(* IEC 61131-3 sources: plc-vscode/tests/st/test-ready/rusty/tests/lit/single/init, 58 files *)

(* ---- array_alias_struct_init.st ---- *)
// RUN: (%COMPILE %s && %RUN) | %CHECK %s

// Verify that array type aliases with struct initializers produce correct runtime values.
TYPE SomeStruct : STRUCT
    field4 : USINT;
END_STRUCT
END_TYPE

TYPE SomeArray : ARRAY[1..2] OF SomeStruct; END_TYPE
TYPE MySomeArrayWInit : SomeArray := [(field4 := 1), (field4 := 2)]; END_TYPE

VAR_GLOBAL
    g_arr : MySomeArrayWInit;
END_VAR

FUNCTION main : DINT
VAR
    local_arr : MySomeArrayWInit;
END_VAR
    // Global instance should carry the type-level initializer
    printf('%d$N', g_arr[1].field4);   // CHECK: 1
    printf('%d$N', g_arr[2].field4);   // CHECK: 2

    // Local instance should also be initialized via the type ctor
    printf('%d$N', local_arr[1].field4);  // CHECK: 1
    printf('%d$N', local_arr[2].field4);  // CHECK: 2
    main := 0;
END_FUNCTION

(* ---- array_constant_indirect_type_init.st ---- *)
// RUN: (%COMPILE %s && %RUN) | %CHECK %s

TYPE IntArrayBase : ARRAY[1..3] OF DINT := [11, 22, 33]; END_TYPE
TYPE IntArrayAlias : IntArrayBase; END_TYPE
TYPE IntArrayAlias2 : IntArrayAlias; END_TYPE

VAR_GLOBAL CONSTANT
    g_base : IntArrayBase;
    g_alias : IntArrayAlias;
    g_alias2 : IntArrayAlias2;
END_VAR

FUNCTION main : DINT
    printf('g_base=%d,%d,%d$N', g_base[1], g_base[2], g_base[3]); // CHECK: g_base=11,22,33
    printf('g_alias=%d,%d,%d$N', g_alias[1], g_alias[2], g_alias[3]); // CHECK: g_alias=11,22,33
    printf('g_alias2=%d,%d,%d$N', g_alias2[1], g_alias2[2], g_alias2[3]); // CHECK: g_alias2=11,22,33

    main := 0;
END_FUNCTION

(* ---- array_external_type_init.st ---- *)
// RUN: (%COMPILE %s && %RUN) | %CHECK %s

// Verify that arrays with type-level initializers work correctly
// when declared in external blocks.
TYPE tarr : ARRAY[0..4] OF DINT := [5(77)]; END_TYPE

VAR_GLOBAL
    g_arr : tarr;
END_VAR

FUNCTION main : DINT
VAR
    local_arr : tarr;
END_VAR
    // Global instance should be initialized by the global ctor
    printf('%d$N', g_arr[0]);   // CHECK: 77
    printf('%d$N', g_arr[4]);   // CHECK: 77

    // Local instance should also be initialized via the type ctor
    printf('%d$N', local_arr[0]);  // CHECK: 77
    printf('%d$N', local_arr[4]);  // CHECK: 77
    main := 0;
END_FUNCTION

(* ---- array_multiplied_large.st ---- *)
// RUN: (%COMPILE %s && %RUN) | %CHECK %s
TYPE tarr : ARRAY[0..9999] OF DINT := [10000(7)]; END_TYPE

FUNCTION main : DINT
VAR
    arr : tarr;
END_VAR
    // Spot-check first, middle, and last elements
    printf('%d$N', arr[0]);     // CHECK: 7
    printf('%d$N', arr[4999]);  // CHECK: 7
    printf('%d$N', arr[9999]);  // CHECK: 7
    main := 0;
END_FUNCTION

(* ---- array_multiplied_mixed_init.st ---- *)
// RUN: (%COMPILE %s && %RUN) | %CHECK %s
TYPE tarr : ARRAY[0..9] OF DINT := [5(10), 3(20), 99, 100]; END_TYPE

FUNCTION main : DINT
VAR
    arr : tarr;
END_VAR
    // First segment: indices 0..4 should be 10
    printf('%d$N', arr[0]);  // CHECK: 10
    printf('%d$N', arr[4]);  // CHECK: 10
    // Second segment: indices 5..7 should be 20
    printf('%d$N', arr[5]);  // CHECK: 20
    printf('%d$N', arr[7]);  // CHECK: 20
    // Individual values at indices 8 and 9
    printf('%d$N', arr[8]);  // CHECK: 99
    printf('%d$N', arr[9]);  // CHECK: 100
    main := 0;
END_FUNCTION

(* ---- array_multiplied_nonzero_offset.st ---- *)
// RUN: (%COMPILE %s && %RUN) | %CHECK %s
TYPE tarr : ARRAY[10..19] OF DINT := [10(77)]; END_TYPE

FUNCTION main : DINT
VAR
    arr : tarr;
END_VAR
    printf('%d$N', arr[10]);  // CHECK: 77
    printf('%d$N', arr[14]);  // CHECK: 77
    printf('%d$N', arr[19]);  // CHECK: 77
    main := 0;
END_FUNCTION

(* ---- array_multiplied_partial_init.st ---- *)
// RUN: (%COMPILE %s && %RUN) | %CHECK %s
TYPE tarr : ARRAY[0..9] OF DINT := [5(42)]; END_TYPE

FUNCTION main : DINT
VAR
    arr : tarr;
END_VAR
    // First 5 elements should be 42
    printf('%d$N', arr[0]);  // CHECK: 42
    printf('%d$N', arr[4]);  // CHECK: 42
    // Remaining elements should be 0 (default)
    printf('%d$N', arr[5]);  // CHECK: 0
    printf('%d$N', arr[9]);  // CHECK: 0
    main := 0;
END_FUNCTION

(* ---- array_multiplied_struct_elements.st ---- *)
// RUN: (%COMPILE %s && %RUN) | %CHECK %s
TYPE MyStruct : STRUCT
    a : DINT;
    b : DINT;
END_STRUCT END_TYPE

FUNCTION main : DINT
VAR
    arr : ARRAY[0..2] OF MyStruct := [3((a := 5, b := 10))];
END_VAR
    printf('%d %d$N', arr[0].a, arr[0].b);  // CHECK: 5 10
    printf('%d %d$N', arr[1].a, arr[1].b);  // CHECK: 5 10
    printf('%d %d$N', arr[2].a, arr[2].b);  // CHECK: 5 10
    main := 0;
END_FUNCTION

(* ---- array_multiplied_type_init.st ---- *)
// RUN: (%COMPILE %s && %RUN) | %CHECK %s
TYPE tarr : ARRAY[0..99] OF DINT := [100(42)]; END_TYPE

FUNCTION main : DINT
VAR
    arr : tarr;
END_VAR
    // Check first, middle, and last elements
    printf('%d$N', arr[0]);   // CHECK: 42
    printf('%d$N', arr[49]);  // CHECK: 42
    printf('%d$N', arr[99]);  // CHECK: 42
    main := 0;
END_FUNCTION

(* ---- array_of_structs_init.st ---- *)
// RUN: (%COMPILE %s && %RUN) | %CHECK %s

TYPE Point : STRUCT
    x : DINT;
    y : DINT;
END_STRUCT END_TYPE

FUNCTION main : DINT
    VAR
        points : ARRAY[0..1] OF Point := [(x := 1, y := 2), (x := 3, y := 4)];
    END_VAR

    // CHECK: 1
    printf('%d$N', points[0].x);

    // CHECK: 2
    printf('%d$N', points[0].y);

    // CHECK: 3
    printf('%d$N', points[1].x);

    // CHECK: 4
    printf('%d$N', points[1].y);
END_FUNCTION

(* ---- global_nested_struct_with_default_and_override_refs.st ---- *)
// RUN: (%COMPILE %s && %RUN) | %CHECK %s
VAR_GLOBAL
    globalValueA: DINT := 5;
    globalValueB: DINT := 10;
    globalValueC: DINT := 15;

    globalStructOne: StructA;
    globalStructTwo: StructA := (value := REF(globalValueA), instanceB := (value := REF(globalValueB), instanceC := (value := REF(globalValueC))));
END_VAR

TYPE StructA:
    STRUCT
        value: REF_TO DINT := REF(globalValueC);
        instanceB: StructB;
    END_STRUCT
END_TYPE

TYPE StructB:
    STRUCT
        value: REF_TO DINT := REF(globalValueA);
        instanceC: StructC;
    END_STRUCT
END_TYPE

TYPE StructC:
    STRUCT
        value: REF_TO DINT := REF(globalValueB);
    END_STRUCT
END_TYPE

FUNCTION main
    printf('%d$N', globalStructOne.value^); // CHECK: 15
    printf('%d$N', globalStructOne.instanceB.value^); // CHECK: 5
    printf('%d$N', globalStructOne.instanceB.instanceC.value^); // CHECK: 10

    printf('%d$N', globalStructTwo.value^); // CHECK: 5
    printf('%d$N', globalStructTwo.instanceB.value^); // CHECK: 10
    printf('%d$N', globalStructTwo.instanceB.instanceC.value^); // CHECK: 15
END_FUNCTION

(* ---- global_nested_struct_with_mixed_ref_assignments.st ---- *)
// RUN: (%COMPILE %s && %RUN) | %CHECK %s
VAR_GLOBAL
    globalOne: DINT := 1;
    globalTwo: DINT := 2;
    globalThree: DINT := 3;
    globalFour: DINT := 4;
    globalFive: DINT := 5;
    globalSix: DINT := 6;
    globalSeven: DINT := 7;
    globalEight: DINT := 8;
    globalNine: DINT := 9;

    globalA: MyStruct2 := (a := (c := REF(globalFive), b := REF(globalSeven)), b := (a := REF(globalThree), b := REF(globalTwo)));
    globalB: MyStruct2 := (b := (a := REF(globalNine)));
END_VAR

TYPE MyStruct2: STRUCT
    a: MyStruct := (a := REF(globalFive), b := REF(globalFour));
    b: MyStruct := (c := REF(globalSeven));
END_STRUCT
END_TYPE

TYPE MyStruct: STRUCT
    a: REF_TO DINT := REF(globalOne);
    b: REF_TO DINT := REF(globalTwo);
    c: REF_TO DINT := REF(globalThree);
END_STRUCT
END_TYPE

FUNCTION main
    printf('%d$N', globalA.a.a^); // CHECK: 5
    printf('%d$N', globalA.a.b^); // CHECK: 7
    printf('%d$N', globalA.a.c^); // CHECK: 5
    printf('%d$N', globalA.b.a^); // CHECK: 3
    printf('%d$N', globalA.b.b^); // CHECK: 2
    printf('%d$N', globalA.b.c^); // CHECK: 7

    printf('%d$N', globalB.b.a^); // CHECK: 9
    printf('%d$N', globalB.b.b^); // CHECK: 2
    printf('%d$N', globalB.b.c^); // CHECK: 7
END_FUNCTION

(* ---- global_struct_with_partial_nested_initialization.st ---- *)
// RUN: (%COMPILE %s && %RUN) | %CHECK %s
VAR_GLOBAL
    globalFoo: DINT := 15;
    globalBar: DINT := 30;
    globalBar2: DINT := 45;

    globalStructOne: StructA;
    globalStructTwo: StructA := (instanceB := (bar := REF(globalBar2)));
END_VAR

TYPE StructA:
    STRUCT
        instanceB: StructB := (foo := REF(globalFoo));
    END_STRUCT
END_TYPE

TYPE StructB:
    STRUCT
        foo: REF_TO DINT;
        bar: REF_TO DINT := REF(globalBar);
    END_STRUCT
END_TYPE

FUNCTION main
    printf('%d$N', globalStructOne.instanceB.foo^); // CHECK: 15
    printf('%d$N', globalStructOne.instanceB.bar^); // CHECK: 30

    printf('%d$N', globalStructTwo.instanceB.foo^); // CHECK: 15
    printf('%d$N', globalStructTwo.instanceB.bar^); // CHECK: 45
END_FUNCTION

(* ---- local_struct_with_global_ref_initialization.st ---- *)
// RUN: (%COMPILE %s && %RUN) | %CHECK %s
VAR_GLOBAL
    globalVar: DINT := 10;
END_VAR

TYPE Parent:
    STRUCT
        foo: REF_TO DINT;
    END_STRUCT
END_TYPE

TYPE Child:
    STRUCT
        instance: Parent := (foo := REF(globalVar));
    END_STRUCT
END_TYPE

FUNCTION main
    VAR
        localChild: Child;
    END_VAR

    // CHECK: Value: 10
    printf('Value: %d$N', localChild.instance.foo^);
END_FUNCTION

(* ---- struct_array_field_init_from_array.st ---- *)
// Issue #921: Array field initialization from another array in struct literal
// RUN: (%COMPILE %s && %RUN) | %CHECK %s

TYPE myStruct : STRUCT
    var1 : DINT;
    var2 : ARRAY[1..2] OF DINT;
END_STRUCT
END_TYPE

FUNCTION main : DINT
VAR
    arr_init : ARRAY[1..2] OF DINT := [1, 2];
    x : myStruct;
END_VAR
    // Initialize array field from another array (regression for #921)
    x := (var1 := 1, var2 := arr_init);

    printf('v1=%d$N', x.var1); // CHECK: v1=1
    printf('v2_1=%d$N', x.var2[1]); // CHECK: v2_1=1
    printf('v2_2=%d$N', x.var2[2]); // CHECK: v2_2=2

    main := 0;
END_FUNCTION

(* ---- struct_with_array_of_strings_init.st ---- *)
// RUN: (%COMPILE %s && %RUN) | %CHECK %s

TYPE Container : STRUCT
    data : ARRAY[0..2] OF STRING;
END_STRUCT END_TYPE

FUNCTION main : DINT
    VAR
        container : Container := (data := ['one', 'two', 'three']);
    END_VAR

    // CHECK: one
    printf('%s$N', container.data[0]);

    // CHECK: two
    printf('%s$N', container.data[1]);

    // CHECK: three
    printf('%s$N', container.data[2]);
END_FUNCTION

(* ---- struct_with_string_init.st ---- *)
// RUN: (%COMPILE %s && %RUN) | %CHECK %s
TYPE Transaction : STRUCT
    id      : DINT;
    amount  : DINT;
    message : STRING;
END_STRUCT END_TYPE

FUNCTION main : DINT
    VAR
        txn     : Transaction := (id := 1, amount := 5, message := 'whats up');
    END_VAR

    // CHECK: 1
    printf('%d$N', txn.id);

    // CHECK: 5
    printf('%d$N', txn.amount);

    // CHECK: whats up
    printf('%s$N', txn.message);
END_FUNCTION

(* ---- type_alias_initializers.st ---- *)
// RUN: (%COMPILE %s && %RUN) | %CHECK %s

// Comprehensive test for type aliases with initializers (enum, struct, array).
TYPE SomeEnum : (E1, E2, E3); END_TYPE
TYPE MySomeEnumWInit : SomeEnum := E2; END_TYPE

TYPE SomeStruct : STRUCT
    field2 : DINT;
    field3 : BOOL;
    field4 : USINT;
END_STRUCT
END_TYPE
TYPE MySomeStructWInit : SomeStruct := (field3 := FALSE, field2 := 9); END_TYPE

TYPE SomeArray : ARRAY[1..2] OF SomeStruct; END_TYPE
TYPE MySomeArrayWInit : SomeArray := [(field4 := 2), (field4 := 2)]; END_TYPE

// Aliases without custom initializers (should inherit defaults)
TYPE MySomeEnum : SomeEnum; END_TYPE
TYPE MySomeStruct : SomeStruct; END_TYPE
TYPE MySomeArray : SomeArray; END_TYPE

FUNCTION main : DINT
VAR
    e : MySomeEnumWInit;
    s : MySomeStructWInit;
    a : MySomeArrayWInit;
    e_default : MySomeEnum;
    s_default : MySomeStruct;
    a_default : MySomeArray;
END_VAR
    // Enum alias with initializer (E1=0, E2=1)
    printf('%d$N', e);            // CHECK: 1

    // Struct alias with initializer
    printf('%d$N', s.field2);     // CHECK: 9
    printf('%d$N', s.field3);     // CHECK: 0

    // Array alias with struct initializer
    printf('%d$N', a[1].field4);  // CHECK: 2
    printf('%d$N', a[2].field4);  // CHECK: 2

    // Default enum (should be 0 / E1)
    printf('%d$N', e_default);    // CHECK: 0

    // Default struct fields (should be 0)
    printf('%d$N', s_default.field2);  // CHECK: 0

    // Default array element (should be 0)
    printf('%d$N', a_default[1].field4);  // CHECK: 0

    main := 0;
END_FUNCTION

(* ---- typedef_initializer_chain.st ---- *)
// Issue #1522: Typedef initializer chains not propagating values
// RUN: (%COMPILE %s && %RUN) | %CHECK %s

TYPE myStruct: STRUCT
  a : INT;
END_STRUCT
END_TYPE

TYPE mytypedefstruct: myStruct := (a := 3); END_TYPE
TYPE mysubtype: mytypedefstruct; END_TYPE
TYPE mysubtype2: mysubtype; END_TYPE

FUNCTION main : DINT
VAR
    inst: mysubtype2;
END_VAR
    printf('a=%d$N', inst.a); // CHECK: a=3
    main := 0;
END_FUNCTION

(* ---- var_input_defaults_function_array_string.st ---- *)
// RUN: (%COMPILE %s && %RUN) | %CHECK %s

// Test VAR_INPUT defaults with STRING/ARRAY and mixed overrides

TYPE ArrType : ARRAY[1..3] OF DINT;
END_TYPE

FUNCTION test : DINT
VAR_INPUT
    s : STRING := 'abc';
    a : ArrType := [1, 2, 3];
END_VAR
test := a[1] + a[2] + a[3];
printf('s=%s$N', REF(s));
printf('sum=%d$N', test);
END_FUNCTION

FUNCTION main
VAR
    tmp : DINT;
END_VAR
// Defaults (no overrides)
tmp := test();
// CHECK: s=abc
// CHECK: sum=6
printf('case=default$N'); // CHECK: case=default

// Override string only
tmp := test(s := 'xyz');
// CHECK: s=xyz
// CHECK: sum=6
printf('case=string$N'); // CHECK: case=string

// Override array only
tmp := test(a := [4, 5, 6]);
// CHECK: s=abc
// CHECK: sum=15
printf('case=array$N'); // CHECK: case=array

// Override both
tmp := test(s := 'pqr', a := [7, 8, 9]);
// CHECK: s=pqr
// CHECK: sum=24
printf('case=both$N'); // CHECK: case=both
END_FUNCTION

(* ---- var_input_defaults_function_wstring.st ---- *)
// RUN: (%COMPILE %s && %RUN) | %CHECK %s
// Test VAR_INPUT defaults with WSTRING and overrides

TYPE ArrType : ARRAY[1..3] OF DINT;
END_TYPE

FUNCTION test : DINT
VAR_INPUT
    s : STRING := 'abc';
    ws : WSTRING := "def";
    a : ArrType := [1, 2, 3];
    i : DINT := 10;
END_VAR
test := a[1] + a[2] + a[3] + i;
printf('s=%s$N', REF(s));
printf('ws=%s$N', REF(TO_STRING(ws)));
printf('sum=%d$N', test);
END_FUNCTION

FUNCTION main : DINT
    // Case 1: all defaults
    test();
    // CHECK: s=abc
    // CHECK: ws=def
    // CHECK: sum=16

    // Case 2: override one input
    test(s := 'xyz');
    // CHECK: s=xyz
    // CHECK: ws=def
    // CHECK: sum=16

    // Case 3: override WSTRING and array
    test(ws := "uvw", a := [4, 5, 6]);
    // CHECK: s=abc
    // CHECK: ws=uvw
    // CHECK: sum=25

    // Case 4: override all inputs
    test(s := 'qqq', ws := "rst", a := [7, 8, 9], i := 1);
    // CHECK: s=qqq
    // CHECK: ws=rst
    // CHECK: sum=25
END_FUNCTION

(* ---- var_input_ref_defaults_string_array.st ---- *)
// RUN: (%COMPILE %s && %RUN) | %CHECK %s
// Test VAR_INPUT {ref} defaults with STRING/ARRAY and mixed overrides

TYPE ArrType : ARRAY[1..3] OF DINT;
END_TYPE

FUNCTION test : DINT
VAR_INPUT {ref}
    s : STRING;
    a : ArrType;
END_VAR
test := a[1] + a[2] + a[3];
printf('s=%s$N', REF(s));
printf('sum=%d$N', test);
END_FUNCTION

FUNCTION main
VAR
    tmp : DINT;
    s_default : STRING := 'abc';
    s_override : STRING := 'xyz';
    s_both : STRING := 'pqr';
    a_default : ArrType := [1, 2, 3];
    a_override : ArrType := [4, 5, 6];
    a_both : ArrType := [7, 8, 9];
END_VAR
// Defaults (no overrides)
tmp := test(s := s_default, a := a_default);
// CHECK: s=abc
// CHECK: sum=6

// Override string only
tmp := test(s := s_override, a := a_default);
// CHECK: s=xyz
// CHECK: sum=6

// Override array only
tmp := test(s := s_default, a := a_override);
// CHECK: s=abc
// CHECK: sum=15

// Override both
tmp := test(s := s_both, a := a_both);
// CHECK: s=pqr
// CHECK: sum=24
END_FUNCTION

(* ---- array_const_bound_multiplied_real.st ---- *)
// RUN: (%COMPILE %s && %RUN) | %CHECK %s
// Tests that an array with constant-expression bounds and a constant-multiplied
// REAL initializer compiles and runs correctly.

VAR_GLOBAL CONSTANT
    NB_BOOL   : DINT := 12;
    NB_ANALOG : DINT := 2;
END_VAR

FUNCTION main : DINT
VAR
    MAX_TIME_BOOL   : ARRAY [1..NB_BOOL] OF REAL := [(NB_BOOL)(0.0033)];
    MAX_TIME_ANALOG : ARRAY [1..NB_ANALOG] OF REAL := [(NB_ANALOG)(1.5)];
END_VAR
    // Check first, middle, and last elements of MAX_TIME_BOOL
    printf('%.4f$N', MAX_TIME_BOOL[1]);   // CHECK: 0.0033
    printf('%.4f$N', MAX_TIME_BOOL[6]);   // CHECK: 0.0033
    printf('%.4f$N', MAX_TIME_BOOL[12]);  // CHECK: 0.0033

    // Check both elements of MAX_TIME_ANALOG
    printf('%.1f$N', MAX_TIME_ANALOG[1]);  // CHECK: 1.5
    printf('%.1f$N', MAX_TIME_ANALOG[2]);  // CHECK: 1.5

    main := 0;
END_FUNCTION

(* ---- array_const_bound_multiplied_real_global.st ---- *)
// RUN: (%COMPILE %s && %RUN) | %CHECK %s
// Tests that global constant arrays with constant-expression bounds and
// constant-multiplied REAL initializers compile and run correctly.

VAR_GLOBAL CONSTANT
    NB_BOOL       : DINT := 12;
    NB_ANALOG     : DINT := 2;
    MAX_TIME_BOOL   : ARRAY [1..NB_BOOL] OF REAL := [(NB_BOOL)(0.0033)];
    MAX_TIME_ANALOG : ARRAY [1..NB_ANALOG] OF REAL := [(NB_ANALOG)(1.5)];
END_VAR

FUNCTION main : DINT
    // Check first, middle, and last elements of MAX_TIME_BOOL
    printf('%.4f$N', MAX_TIME_BOOL[1]);   // CHECK: 0.0033
    printf('%.4f$N', MAX_TIME_BOOL[6]);   // CHECK: 0.0033
    printf('%.4f$N', MAX_TIME_BOOL[12]);  // CHECK: 0.0033

    // Check both elements of MAX_TIME_ANALOG
    printf('%.1f$N', MAX_TIME_ANALOG[1]);  // CHECK: 1.5
    printf('%.1f$N', MAX_TIME_ANALOG[2]);  // CHECK: 1.5

    main := 0;
END_FUNCTION

(* ---- global_variables.st ---- *)
// RUN: (%COMPILE %s && %RUN) | %CHECK %s
VAR_GLOBAL
    arr : ARRAY[0..3] OF STRING := ['a', 'b', 'c', 'd'];
    alias AT arr : ARRAY[0..3] OF STRING;
END_VAR

FUNCTION main: DINT
    // CHECK: a, b, c, d
    printf('%s, %s, %s, %s$N', REF(alias[0]), REF(alias[1]), REF(alias[2]), REF(alias[3]));
END_FUNCTION

(* ---- ref_initializer_with_array_init.st ---- *)
// RUN: (%COMPILE %s && %RUN) | %CHECK %s

VAR_GLOBAL
    globalString: STRING := 'Global String';
END_VAR

FUNCTION main : DINT
VAR
    localString: REF_TO STRING := REF(globalString);
    arr: ARRAY[1..2] OF DINT := [1, 2];
END_VAR
    printf('ref=%s$N', localString); // CHECK: ref=Global String
    printf('arr1=%d$N', arr[1]); // CHECK: arr1=1
    printf('arr2=%d$N', arr[2]); // CHECK: arr2=2
    main := 0;
END_FUNCTION

(* ---- array_local_const_multiplied.st ---- *)
// RUN: (%COMPILE %s && %RUN) | %CHECK %s
// Tests that a POU-local VAR CONSTANT can be used as the multiplier
// in an array initializer with the [(CONST)(value)] syntax.

FUNCTION main : DINT
VAR CONSTANT
    N     : DINT := 5;
    COUNT : DINT := 3;
END_VAR
VAR
    arr1 : ARRAY [0..4] OF DINT := [(N)(77)];
    arr2 : ARRAY [1..3] OF REAL := [(COUNT)(1.25)];
END_VAR
    printf('%d$N', arr1[0]);  // CHECK: 77
    printf('%d$N', arr1[2]);  // CHECK: 77
    printf('%d$N', arr1[4]);  // CHECK: 77

    printf('%.2f$N', arr2[1]);  // CHECK: 1.25
    printf('%.2f$N', arr2[3]);  // CHECK: 1.25

    main := 0;
END_FUNCTION

(* ---- array_mixed_ref_segments.st ---- *)
// RUN: (%COMPILE %s && %RUN) | %CHECK %s
// Tests mixed multiplied segments with REF() calls.
FUNCTION main : DINT
VAR
    a : DINT := 1;
    b : DINT := 2;
    arr : ARRAY[0..4] OF REF_TO DINT := [2(REF(a)), REF(b), 2(REF(a))];
END_VAR
    printf('%d$N', arr[0]^);  // CHECK: 1
    printf('%d$N', arr[1]^);  // CHECK: 1
    printf('%d$N', arr[2]^);  // CHECK: 2
    printf('%d$N', arr[3]^);  // CHECK: 1
    printf('%d$N', arr[4]^);  // CHECK: 1
    main := 0;
END_FUNCTION

(* ---- array_multiplied_initializer_with_variable.st ---- *)
// RUN: (%COMPILE %s && %RUN) | %CHECK %s
FUNCTION main : INT
    VAR
        arr : ARRAY[1..32] OF INT := [32(1)];
        x : INT;
    END_VAR

    x := 5;
    arr := [32(x)];

    // CHECK: 15
    printf('%d$N', arr[1] + arr[16] + arr[32]);
END_FUNCTION

(* ---- array_of_strings_init.st ---- *)
// RUN: (%COMPILE %s && %RUN) | %CHECK %s

FUNCTION main : DINT
    VAR
        arr : ARRAY[0..2] OF STRING := ['apple', 'banana', 'cherry'];
    END_VAR

    // CHECK: apple
    printf('%s$N', arr[0]);

    // CHECK: banana
    printf('%s$N', arr[1]);

    // CHECK: cherry
    printf('%s$N', arr[2]);
END_FUNCTION

(* ---- array_ref_elements.st ---- *)
// RUN: (%COMPILE %s && %RUN) | %CHECK %s
// Tests that arrays initialized with REF() (runtime function calls) are
// correctly lowered into indexed assignments.
FUNCTION main : DINT
VAR
    a : DINT := 10;
    b : DINT := 20;
    c : DINT := 30;
    arr_mult : ARRAY[0..2] OF REF_TO DINT := [3(REF(a))];
    arr_list : ARRAY[0..2] OF REF_TO DINT := [REF(a), REF(b), REF(c)];
END_VAR
    // Multiplied: all point to a
    printf('%d$N', arr_mult[0]^);  // CHECK: 10
    printf('%d$N', arr_mult[1]^);  // CHECK: 10
    printf('%d$N', arr_mult[2]^);  // CHECK: 10

    // Expression list: each points to a different variable
    printf('%d$N', arr_list[0]^);  // CHECK: 10
    printf('%d$N', arr_list[1]^);  // CHECK: 20
    printf('%d$N', arr_list[2]^);  // CHECK: 30

    // Verify they are actual pointers (mutation through ref)
    arr_list[1]^ := 99;
    printf('%d$N', b);  // CHECK: 99
    main := 0;
END_FUNCTION

(* ---- array_variable_elements.st ---- *)
// RUN: (%COMPILE %s && %RUN) | %CHECK %s
// Tests that arrays initialized with variable references (non-constant
// expressions) are correctly lowered into indexed assignments.
FUNCTION main : DINT
VAR
    x : DINT := 42;
    y : DINT := 7;
    arr_mult : ARRAY[0..2] OF DINT := [3(x)];
    arr_list : ARRAY[0..3] OF DINT := [x, y, x, y];
END_VAR
    // Multiplied: all get value of x at init time
    printf('%d$N', arr_mult[0]);  // CHECK: 42
    printf('%d$N', arr_mult[1]);  // CHECK: 42
    printf('%d$N', arr_mult[2]);  // CHECK: 42

    // Expression list: alternating x and y
    printf('%d$N', arr_list[0]);  // CHECK: 42
    printf('%d$N', arr_list[1]);  // CHECK: 7
    printf('%d$N', arr_list[2]);  // CHECK: 42
    printf('%d$N', arr_list[3]);  // CHECK: 7
    main := 0;
END_FUNCTION

(* ---- var_inout_not_initialized.st ---- *)
// RUN: (%COMPILE %s && %RUN) | %CHECK %s
// Test that VAR_IN_OUT parameters without initializers keep their passed values
// Note: VAR_IN_OUT initializers are NOT applied in the current implementation

FUNCTION test_no_init
VAR_IN_OUT
    value : INT;
END_VAR
    // CHECK: 42
    printf('%d$N', value);
END_FUNCTION

FUNCTION main: DINT
    VAR
        x : INT;
    END_VAR
    x := 42;
    test_no_init(x);
END_FUNCTION

(* ---- config_variables.st ---- *)
// RUN: (%COMPILE %s && %RUN) | %CHECK %s
FUNCTION_BLOCK FB
VAR
  foo AT %I* : DINT;
END_VAR
    printf('%d$N', foo);
END_FUNCTION_BLOCK

VAR_CONFIG
  prog.instance1.foo AT %IX1.2.1 : DINT;
  prog.instance2.foo AT %QX1.2.2 : DINT;
END_VAR

PROGRAM prog
VAR
    instance1: FB;
    instance2: FB;
END_VAR
    instance1(); // CHECK: 23
    instance2(); // CHECK: 48
END_PROGRAM

FUNCTION main : DINT
    %IX1.2.1 := 23;
    %QX1.2.2 := 48;
    prog();
END_FUNCTION

(* ---- config_variables_dont_clash_with_globals.st ---- *)
// RUN: (%COMPILE %s && %RUN) | %CHECK %s
FUNCTION_BLOCK FB
VAR
  foo AT %I* : DINT;
END_VAR
    printf('%d$N', foo);
END_FUNCTION_BLOCK

VAR_CONFIG
  prog.instance1.foo AT %IX1.2.1 : DINT;
  prog.instance2.foo AT %QX1.2.2 : DINT;
END_VAR

VAR_GLOBAL
    a AT %IX1.2.1 : DINT;
    b AT %QX1.2.2 : DINT;
END_VAR

PROGRAM prog
VAR
    instance1: FB;
    instance2: FB;
END_VAR
    instance1(); // CHECK: 23
    instance2(); // CHECK: 48
END_PROGRAM

FUNCTION main : DINT
    a := 23;
    b := 48;
    prog();
END_FUNCTION

(* ---- function_locals.st ---- *)
// RUN: (%COMPILE %s && %RUN) | %CHECK %s
VAR_GLOBAL
    ps: STRING := 'Hello world!';
    ps2: STRING;
    x : DINT := 1337;
END_VAR

FUNCTION_BLOCK foo
VAR
    s AT ps: STRING;
END_VAR
VAR_TEMP
    s2 AT ps2: STRING;
END_VAR
    s2 := 'Hello from me, too';

    // CHECK: Hello world!
    printf('%s$N', REF(s));
    // CHECK: Hello from me, too
    printf('%s$N', REF(s2));
END_FUNCTION_BLOCK

FUNCTION_BLOCK bar
VAR
    x : DINT := 69;
    shadowed_global : REF_TO DINT := REF(x);
    alias_to_local AT x : DINT;
    reference_to_local : REFERENCE TO DINT REF= x;
END_VAR
VAR_TEMP
    y : DINT := 420;
    temp_ref_to_temp : REF_TO DINT := REF(y);
    temp_alias AT y :DINT;
    temp_reference_to : REFERENCE TO DINT REF= y;
END_VAR
    printf('%d$N', shadowed_global^); // CHECK: 69
    printf('%d$N', temp_ref_to_temp^); // CHECK: 420
    printf('%d$N', alias_to_local); // CHECK: 69
    printf('%d$N', reference_to_local); // CHECK: 69
    printf('%d$N', temp_alias); // CHECK: 420
    printf('%d$N', temp_reference_to); // CHECK: 420
END_FUNCTION_BLOCK

FUNCTION main: DINT
VAR
    fb: foo;
    bb: bar;

    z : DINT := 42;
    temp_ref_to_temp : REF_TO DINT := REF(z);
    temp_alias AT z :DINT;
    temp_reference_to : REFERENCE TO DINT REF= z;
END_VAR
    fb();
    bb();

    printf('%d$N', temp_ref_to_temp^); // CHECK: 42
    printf('%d$N', temp_alias); // CHECK: 42
    printf('%d$N', temp_reference_to); // CHECK: 42

    baz();
END_FUNCTION

FUNCTION baz
    VAR
        s1: REF_TO LINT := REF(t1);
        s2 AT t1 : LINT;
        s3 : REFERENCE TO LINT REF= t1;
        s4 AT s2 : LINT;
        s5 : REF_TO LINT := REF(s4);
        s6 : REFERENCE TO LINT REF= s4;
    END_VAR
    VAR_TEMP
        t1 : LINT := 16#DEADBEEF;
        t2 : REF_TO LINT := REF(t1);
        t3 AT s2 : LINT;
        t4 : REFERENCE TO LINT REF= s4;
    END_VAR
        printf('%#010x$N', s1^);    // CHECK: 0xdeadbeef
        printf('%#010x$N', s2);     // CHECK: 0xdeadbeef
        printf('%#010x$N', s3);     // CHECK: 0xdeadbeef
        printf('%#010x$N', s4);     // CHECK: 0xdeadbeef
        printf('%#010x$N', s5^);    // CHECK: 0xdeadbeef
        printf('%#010x$N', s6);     // CHECK: 0xdeadbeef
        printf('%#010x$N', t2^);    // CHECK: 0xdeadbeef
        printf('%#010x$N', t3);     // CHECK: 0xdeadbeef
        printf('%#010x$N', t4);     // CHECK: 0xdeadbeef
END_FUNCTION

(* ---- global_struct_instances.st ---- *)
// RUN: (%COMPILE %s && %RUN) | %CHECK %s
VAR_GLOBAL
    arr : ARRAY[1..3] OF DINT := [3, 2, 1];
    foo: foo_t;
END_VAR

FUNCTION_BLOCK foo_t
VAR
    refArr AT arr : ARRAY[1..3] OF DINT;
END_VAR
    // CHECK: 1, 2, 3
    printf('%d, %d, %d$N', refArr[3], refArr[2], refArr[1]);
END_FUNCTION_BLOCK

FUNCTION main: DINT
    foo();
END_FUNCTION

(* ---- methods.st ---- *)
// RUN: (%COMPILE %s && %RUN) | %CHECK %s
VAR_GLOBAL CONSTANT
    g2 : STRING := 'Whats up';
END_VAR

VAR_GLOBAL
    g0 : DINT := 5;

    // g1 used to be a constant in this test, but now we have explicit validation that says that constants cannot be referenced in pointers
    g1 : Transaction := (id := 5, amount := 10, message := g2);
END_VAR

TYPE Transaction : STRUCT
    id      : DINT;
    amount  : DINT;
    message : STRING;
END_STRUCT END_TYPE

FUNCTION_BLOCK fb0
VAR
    s : STRING := 'hello from foo';
END_VAR
    METHOD fbMethod
        VAR
            local_s AT s: STRING;
        END_VAR
        VAR_TEMP
            local_s2 AT local_s: STRING;
            ptr : REF_TO STRING := REF(local_s2);
        END_VAR
            // CHECK: hello from foo
            printf('%s$N', ptr);
    END_METHOD
END_FUNCTION_BLOCK

FUNCTION_BLOCK fb1
    VAR
        foo : DINT := 5;
    END_VAR

    METHOD fbMethod
        VAR
            bar : REFERENCE TO DINT := REF(foo);
        END_VAR

        printf('%d$N', bar); // CHECK: 5
    END_METHOD
END_FUNCTION_BLOCK

FUNCTION_BLOCK fb2
    VAR
        foo AT g0 : DINT;
    END_VAR

    METHOD fbMethod
        VAR
            bar : REFERENCE TO DINT := REF(baz);
            baz : REFERENCE TO DINT := REF(foo);
        END_VAR

        printf('%d$N', baz); // CHECK: 5
    END_METHOD
END_FUNCTION_BLOCK

FUNCTION_BLOCK fb3
    VAR
        foo : DINT := 5;
    END_VAR

    METHOD fbMethod
        VAR
            bar : REFERENCE TO DINT := REF(baz);
            baz : REFERENCE TO DINT := REF(foo);
        END_VAR

        printf('%d$N', baz); // CHECK: 5
    END_METHOD
END_FUNCTION_BLOCK

FUNCTION_BLOCK fb4
    VAR
        foo : Transaction := (id := 5, amount := 10, message := 'Whats up');
    END_VAR

    METHOD fbMethod
        VAR
            bar : REFERENCE TO Transaction := REF(baz);
            baz : REFERENCE TO Transaction := REF(foo);
        END_VAR

        printf('%d$N', foo.id);         // CHECK: 5
        printf('%d$N', foo.amount);     // CHECK: 10
        printf('%s$N', REF(foo.message));    // CHECK: Whats up
    END_METHOD
END_FUNCTION_BLOCK

FUNCTION_BLOCK fb5
    METHOD fbMethod
        VAR
            bar : REFERENCE TO DINT := REF(g0);
        END_VAR

        printf('%d$N', bar); // CHECK: 5
    END_METHOD
END_FUNCTION_BLOCK

FUNCTION_BLOCK fb6
    METHOD fbMethod
        VAR
            bar : REFERENCE TO Transaction := REF(g1);
        END_VAR

        printf('%d$N', g1.id);         // CHECK: 5
        printf('%d$N', g1.amount);     // CHECK: 10
        printf('%s$N', REF(g1.message));    // CHECK: Whats up
    END_METHOD
END_FUNCTION_BLOCK

PROGRAM prog
    VAR
        fb0: fb0;
        fb1: fb1;
        fb2: fb2;
        fb3: fb3;
    END_VAR
    METHOD progMethod
        VAR
            fb4: fb4;
            fb5: fb5;
            fb6: fb6;
        END_VAR
            fb0.fbMethod();
            fb1.fbMethod();
            fb2.fbMethod();
            fb3.fbMethod();
            fb4.fbMethod();
            fb5.fbMethod();
            fb6.fbMethod();
    END_METHOD
    progMethod();
END_PROGRAM

FUNCTION main : DINT
VAR
    fb0: fb0;
    fb1: fb1;
    fb2: fb2;
    fb3: fb3;
    fb4: fb4;
    fb5: fb5;
    fb6: fb6;
END_VAR
    fb0.fbMethod();
    fb1.fbMethod();
    fb2.fbMethod();
    fb3.fbMethod();
    fb4.fbMethod();
    fb5.fbMethod();
    fb6.fbMethod();
    prog();
END_FUNCTION

(* ---- nested_pous.st ---- *)
// RUN: (%COMPILE %s && %RUN) | %CHECK %s
VAR_GLOBAL
    arr : ARRAY[1..3] OF DINT;
END_VAR

FUNCTION_BLOCK foo_t
VAR
    refArr AT arr : ARRAY[1..3] OF DINT;
END_VAR
    arr[1] := 3;
    arr[2] := 2;
    arr[3] := 1;

    // CHECK: 1, 2, 3
    printf('%d, %d, %d$N', refArr[3], refArr[2], refArr[1]);
END_FUNCTION_BLOCK

FUNCTION_BLOCK bar_t
VAR
    foo: foo_t;
END_VAR
    foo();
END_FUNCTION_BLOCK

PROGRAM baz
VAR
    refArr AT arr : ARRAY[1..3] OF DINT;
    bar: bar_t;
END_VAR
    arr[1] := 3;
    arr[2] := 2;
    arr[3] := 1;

    // CHECK: 1, 2, 3
    printf('%d, %d, %d$N', refArr[3], refArr[2], refArr[1]);

    bar();
END_PROGRAM

FUNCTION main: DINT
    baz();
END_FUNCTION

(* ---- ref_override_in_initializer.st ---- *)
// RUN: (%COMPILE %s && %RUN) | %CHECK %s

VAR_GLOBAL
    ps: INT := 42;
END_VAR

PROGRAM mainProg
VAR
    fb: foo := (s1 := REF(ps));
END_VAR
END_PROGRAM

FUNCTION_BLOCK foo
VAR
    default_target: INT := 11;
END_VAR
VAR_INPUT
    s1: REF_TO INT := REF(default_target);
END_VAR

METHOD get_value : INT
    get_value := s1^;
END_METHOD

METHOD set_value
VAR_INPUT
    v: INT;
END_VAR
    s1^ := v;
END_METHOD
END_FUNCTION_BLOCK

FUNCTION main
VAR
    out_val: INT;
END_VAR
    out_val := mainProg.fb.get_value();
    printf('read_from_ref=%d$N', out_val); // CHECK: read_from_ref=42

    mainProg.fb.set_value(v := 77);
    printf('write_via_ref=%d$N', ps); // CHECK: write_via_ref=77
END_FUNCTION

(* ---- struct_literal_local_qualifier.st ---- *)
// RUN: (%COMPILE %s && %RUN) | %CHECK %s

TYPE MyStruct : STRUCT
    field : DINT;
END_STRUCT
END_TYPE

VAR_GLOBAL
    local : DINT := 5;
END_VAR

FUNCTION_BLOCK Foo
VAR
    local : DINT := 42;
    s : MyStruct := (field := local);
END_VAR
END_FUNCTION_BLOCK

PROGRAM prog
VAR
    fb : Foo;
END_VAR
    // CHECK: 42
    printf('%d$N', fb.s.field);
END_PROGRAM

FUNCTION main : DINT
    prog();
END_FUNCTION

(* ---- struct_with_fb_member.st ---- *)
// RUN: (%COMPILE %s && %RUN) | %CHECK %s

TYPE MyStruct : STRUCT
    fb : FbA := (x := 10);
END_STRUCT
END_TYPE

FUNCTION_BLOCK FbA
VAR
    x : DINT;
END_VAR
END_FUNCTION_BLOCK

FUNCTION main : DINT
VAR
    s : MyStruct;
END_VAR
    // CHECK: s.fb.x = 10
    printf('s.fb.x = %d$N', s.fb.x);
END_FUNCTION

(* ---- user_init.st ---- *)
// RUN: (%COMPILE %s && %RUN) | %CHECK %s
TYPE
    bar : STRUCT
        f: foo;
    END_STRUCT;
END_TYPE

FUNCTION_BLOCK foo
VAR
    x : INT := 0;
    y : INT := 0;
END_VAR
    METHOD FB_INIT
        x := 1;
        y := 2;
    END_METHOD
END_FUNCTION_BLOCK

PROGRAM prog
VAR
    str: bar;
END_VAR
    printf('%d$N', str.f.x); // CHECK: 1
    printf('%d$N', str.f.y); // CHECK: 2
END_PROGRAM

FUNCTION main: DINT
    prog();
END_FUNCTION

(* ---- user_init_for_stack_variable.st ---- *)
// RUN: (%COMPILE %s && %RUN) | %CHECK %s
FUNCTION_BLOCK foo
    METHOD FB_INIT
        printf('FB_INIT called$N');
    END_METHOD
END_FUNCTION_BLOCK

FUNCTION main
VAR
    fb: foo;
END_VAR
    // CHECK: FB_INIT called
END_FUNCTION

(* ---- array_assignment_in_body.st ---- *)
// Test to verify array assignment works in body (not initializer)
// This test confirms that array assignment works correctly when done in the body
// rather than as an initializer, which helps isolate initializer-specific issues.
// RUN: (%COMPILE %s && %RUN) | %CHECK %s

VAR_GLOBAL
    g1: INT := 10;
    g2: INT := 20;
END_VAR

TYPE Elem: STRUCT
    r: REF_TO INT := REF(g1);
END_STRUCT END_TYPE

PROGRAM mainProg
VAR
    arr: ARRAY[1..2] OF Elem;
END_VAR
    // Assign array in one go
    arr := [
        (r := REF(g1)),
        (r := REF(g2))
    ];
END_PROGRAM

FUNCTION main : DINT
VAR
    v1: INT;
    v2: INT;
END_VAR
    mainProg();
    v1 := mainProg.arr[1].r^;
    v2 := mainProg.arr[2].r^;
    printf('v1=%d$N', v1); // CHECK: v1=10
    printf('v2=%d$N', v2); // CHECK: v2=20
    mainProg.arr[1].r^ := 33;
    mainProg.arr[2].r^ := 44;
    printf('g1=%d$N', g1); // CHECK: g1=33
    printf('g2=%d$N', g2); // CHECK: g2=44
    main := 0;
END_FUNCTION

(* ---- array_multidim_and_nested_init.st ---- *)
// RUN: (%COMPILE %s && %RUN) | %CHECK %s
// Tests initialization of multi-dimensional arrays and arrays of arrays,
// including struct element types.

TYPE str1 : STRUCT
    a : INT;
END_STRUCT END_TYPE

PROGRAM mainProg
VAR
    x2 : ARRAY [0..1, 0..1] OF INT := [11,12,21,22];
    x3 : ARRAY [0..1] OF ARRAY[0..1] OF INT := [[11,12],[21,22]];

    x2_1 : ARRAY [0..1, 0..1] OF str1 := [(a:=11),(a:=12),(a:=21),(a:=22)];
    x3_1 : ARRAY [0..1] OF ARRAY[0..1] OF str1 := [[(a:=11),(a:=12)],[(a:=21),(a:=22)]];
END_VAR
    ;
END_PROGRAM

FUNCTION main : DINT
    mainProg();

    // Multi-dimensional array of INT
    // CHECK: x2=11,12,21,22
    printf('x2=%d,%d,%d,%d$N', mainProg.x2[0,0], mainProg.x2[0,1], mainProg.x2[1,0], mainProg.x2[1,1]);

    // Array of array of INT
    // CHECK: x3=11,12,21,22
    printf('x3=%d,%d,%d,%d$N', mainProg.x3[0][0], mainProg.x3[0][1], mainProg.x3[1][0], mainProg.x3[1][1]);

    // Multi-dimensional array of struct
    // CHECK: x2_1=11,12,21,22
    printf('x2_1=%d,%d,%d,%d$N', mainProg.x2_1[0,0].a, mainProg.x2_1[0,1].a, mainProg.x2_1[1,0].a, mainProg.x2_1[1,1].a);

    // Array of array of struct
    // CHECK: x3_1=11,12,21,22
    printf('x3_1=%d,%d,%d,%d$N', mainProg.x3_1[0][0].a, mainProg.x3_1[0][1].a, mainProg.x3_1[1][0].a, mainProg.x3_1[1][1].a);

    main := 0;
END_FUNCTION

(* ---- array_multiplied_variable_override.st ---- *)
// RUN: (%COMPILE %s && %RUN) | %CHECK %s
TYPE tarr : ARRAY[0..9] OF DINT := [10(42)]; END_TYPE

PROGRAM prog
VAR
    default_arr : tarr;
    override_arr : tarr := [10(99)];
END_VAR
    printf('%d$N', default_arr[0]);   // CHECK: 42
    printf('%d$N', default_arr[9]);   // CHECK: 42
    printf('%d$N', override_arr[0]);  // CHECK: 99
    printf('%d$N', override_arr[9]);  // CHECK: 99
END_PROGRAM

FUNCTION main : DINT
    prog();
    main := 0;
END_FUNCTION

(* ---- array_partial_init_warning.st ---- *)
// RUN: (%COMPILE %s && %RUN) | %CHECK %s
// Tests that partial array initialization zero-pads at runtime.

PROGRAM mainProg
VAR
    a1 : ARRAY [0..3] OF INT := [10, 20];
    a2 : ARRAY [0..1, 0..1] OF INT := [10, 20, 30];
    a3 : ARRAY [0..1] OF ARRAY[0..1] OF INT := [[10, 20]];
END_VAR
    ;
END_PROGRAM

FUNCTION main : DINT
    mainProg();

    // CHECK: a1=10,20,0,0
    printf('a1=%d,%d,%d,%d$N', mainProg.a1[0], mainProg.a1[1], mainProg.a1[2], mainProg.a1[3]);

    // CHECK: a2=10,20,30,0
    printf('a2=%d,%d,%d,%d$N', mainProg.a2[0,0], mainProg.a2[0,1], mainProg.a2[1,0], mainProg.a2[1,1]);

    // CHECK: a3=10,20,0,0
    printf('a3=%d,%d,%d,%d$N', mainProg.a3[0][0], mainProg.a3[0][1], mainProg.a3[1][0], mainProg.a3[1][1]);

    main := 0;
END_FUNCTION

(* ---- array_partial_init_warning_type_and_var.st ---- *)
// RUN: not %PLC --check --error-format clang --error-config %S/../../util/diagnostics_e127_as_error.json %s 2>&1 | %CHECK %s
// E127 is promoted to error so we can assert both diagnostics are emitted.
// CHECK-DAG: {{.*}}array_partial_init_warning_type_and_var.st:{{[0-9]+}}:{{[0-9]+}}:{{.*}}error[E127]: Fewer initial values for array `a` than expected. Expected 5, found 2.
// CHECK-DAG: {{.*}}array_partial_init_warning_type_and_var.st:{{[0-9]+}}:{{[0-9]+}}:{{.*}}error[E127]: Fewer initial values for array `userArrayType` than expected. Expected 5, found 4.

PROGRAM PLC_PRG
    VAR CONSTANT
        x : INT := 0;
    END_VAR
    VAR
        a : userArrayType := [x,x];
    END_VAR
END_PROGRAM

TYPE userArrayType : ARRAY [1..5] OF INT := [1,2,4,5];
END_TYPE

(* ---- array_single_element_init.st ---- *)
// RUN: (%COMPILE %s && %RUN) | %CHECK %s
// Tests that single-element array initialization compiles and zero-pads correctly.

PROGRAM mainProg
VAR
    a1 : ARRAY [0..3] OF INT := [11];
    a2 : ARRAY [0..1, 0..1] OF INT := [42];
    a3 : ARRAY [0..1] OF ARRAY[0..1] OF INT := [[99]];
END_VAR
    ;
END_PROGRAM

FUNCTION main : DINT
    mainProg();

    // 1D: first element set, rest zero
    // CHECK: a1=11,0,0,0
    printf('a1=%d,%d,%d,%d$N', mainProg.a1[0], mainProg.a1[1], mainProg.a1[2], mainProg.a1[3]);

    // 2D flat: first element set, rest zero
    // CHECK: a2=42,0,0,0
    printf('a2=%d,%d,%d,%d$N', mainProg.a2[0,0], mainProg.a2[0,1], mainProg.a2[1,0], mainProg.a2[1,1]);

    // Nested: first inner element set, rest zero
    // CHECK: a3=99,0,0,0
    printf('a3=%d,%d,%d,%d$N', mainProg.a3[0][0], mainProg.a3[0][1], mainProg.a3[1][0], mainProg.a3[1][1]);

    main := 0;
END_FUNCTION

(* ---- array_struct_ref_initialization.st ---- *)
// Issue #1295: Array of structs with ref-initialized fields
// RUN: (%COMPILE %s && %RUN) | %CHECK %s

VAR_GLOBAL
    g1: INT := 10;
    g2: INT := 20;
END_VAR

TYPE Elem: STRUCT
    r: REF_TO INT := REF(g1);
END_STRUCT END_TYPE

PROGRAM mainProg
VAR
    arr: ARRAY[1..2] OF Elem := [
        (r := REF(g1)),
        (r := REF(g2))
    ];
END_VAR
END_PROGRAM

FUNCTION main : DINT
VAR
    v1: INT;
    v2: INT;
END_VAR
    v1 := mainProg.arr[1].r^;
    v2 := mainProg.arr[2].r^;
    printf('v1=%d$N', v1); // CHECK: v1=10
    printf('v2=%d$N', v2); // CHECK: v2=20
    mainProg.arr[1].r^ := 33;
    mainProg.arr[2].r^ := 44;
    printf('g1=%d$N', g1); // CHECK: g1=33
    printf('g2=%d$N', g2); // CHECK: g2=44
    main := 0;
END_FUNCTION

(* ---- mixed_parameter_types_with_structs.st ---- *)
// RUN: (%COMPILE %s && %RUN) | %CHECK %s
// Test mixed VAR_INPUT and VAR_IN_OUT parameters

FUNCTION test_mixed_params
VAR_INPUT
    input_val : INT;
    input_str : STRING;
END_VAR
VAR_IN_OUT
    inout_val : INT;
END_VAR
    // CHECK: 5
    printf('%d$N', input_val);

    // CHECK: hello
    printf('%s$N', input_str);

    // CHECK: 42
    printf('%d$N', inout_val);
END_FUNCTION

PROGRAM prog
VAR
    x : INT;
END_VAR
    x := 42;
    test_mixed_params(5, 'hello', x);
END_PROGRAM

FUNCTION main: DINT
    prog();
END_FUNCTION

(* ---- program.st ---- *)
// RUN: (%COMPILE %s && %RUN) | %CHECK %s
VAR_GLOBAL
    gs: STRING;
END_VAR

PROGRAM prog
VAR
    s AT gs: STRING;
END_VAR
    s := 'Hello world!';

    // CHECK: Hello world!
    printf('%s$N', REF(gs));
END_PROGRAM

FUNCTION main: DINT
    prog();
END_FUNCTION

(* ---- struct_ref_literal_paren.st ---- *)
// RUN: (%COMPILE %s && %RUN) | %CHECK %s

VAR_GLOBAL
    g : DINT := 21;
END_VAR

TYPE MyStruct : STRUCT
    r : REFERENCE TO DINT;
END_STRUCT
END_TYPE

VAR_GLOBAL
    s : MyStruct := (r := (REF(g)));
END_VAR

PROGRAM prog
    // CHECK: 21
    printf('%d$N', s.r);
END_PROGRAM

FUNCTION main : DINT
    prog();
END_FUNCTION

(* ---- structs.st ---- *)
// RUN: (%COMPILE %s && %RUN) | %CHECK %s
VAR_GLOBAL CONSTANT
    constantDintValue : DINT := 12345;
END_VAR
TYPE myStruct : STRUCT
        member : REF_TO STRING := REF(s);
        member2 AT s2 : ARRAY[0..1] OF STRING;
        member3: DINT := 367;
        member4: DINT := 12345;
    END_STRUCT
END_TYPE

VAR_GLOBAL
    s : STRING := 'Hello, world!';
    s2 : ARRAY[0..1] OF STRING := ['hello', 'world'];
END_VAR

PROGRAM prog
VAR
    str: myStruct;
END_VAR
VAR_TEMP
    tmp: STRING;
END_VAR
    // CHECK: Hello, world!
    printf('%s$N', str.member);
    // CHECK: hello world
    tmp := str.member2[0];
    printf('%s', REF(tmp));
    tmp := str.member2[1];
    printf(' %s$N', REF(tmp));
    // CHECK: 367
    printf('%d$N', str.member3);
    // CHECK: 12345
    printf('%d$N', str.member4);
END_PROGRAM

FUNCTION main: DINT
    prog();
END_FUNCTION

(* ---- var_inout_with_init_stack_constructor.st ---- *)
// RUN: (%COMPILE %s && %RUN) | %CHECK %s
// Test that VAR_IN_OUT with initializers keeps passed values

FUNCTION test_inout_no_init
VAR_IN_OUT
    x : INT;
END_VAR
    // CHECK: 42
    printf('%d$N', x);
END_FUNCTION

PROGRAM prog
VAR
    v : INT;
END_VAR
    v := 42;
    test_inout_no_init(v);
END_PROGRAM

FUNCTION main: DINT
    prog();
END_FUNCTION

(* ---- var_input_with_init.st ---- *)
// RUN: (%COMPILE %s && %RUN) | %CHECK %s
// Test that VAR_INPUT variables can be initialized

PROGRAM TestVarInput
VAR_INPUT
    x : INT := 42;
    s : STRING := 'hello';
END_VAR
VAR
    result : INT;
END_VAR
    result := x;

    // CHECK: 42
    printf('%d$N', result);

    // CHECK: hello
    printf('%s$N', s);
END_PROGRAM

FUNCTION main: DINT
    TestVarInput();
END_FUNCTION

(* ---- var_output_with_init.st ---- *)
// RUN: (%COMPILE %s && %RUN) | %CHECK %s
// Test that VAR_OUTPUT variables can be initialized

PROGRAM TestVarOutput
VAR_OUTPUT
    result : INT := 99;
    msg : STRING := 'output';
END_VAR

    // CHECK: 99
    printf('%d$N', result);

    // CHECK: output
    printf('%s$N', msg);
END_PROGRAM

FUNCTION main: DINT
    TestVarOutput();
END_FUNCTION
